// TIA Portal V21 export
// export: Created 2026-11-11T00:47:22.4274178Z, ExportSetting WithDefaults, DisplayName Totally Integrated Automation Portal, DisplayVersion V21 Update 3, DisplayName STEP 7 Professional, DisplayVersion V21 Update 3, DisplayName STEP 7 Safety, DisplayVersion V21, DisplayName Tech WebApplication, DisplayVersion V21, DisplayName WinCC Basic/Comfort/Advanced, DisplayVersion V21 Update 3, DisplayName WinCC Unified, DisplayVersion V21 Update 3
FUNCTION_BLOCK "FB_Fbd_ex066"   // FB102, FBD
{ S7_Optimized_Access := 'TRUE' }
VERSION : 0.1
// stored: AutoNumber true, IsIECCheckEnabled false, IsRetainMemResEnabled false, MemoryReserve 100, SetENOAutomatically false, UDAEnableTagReadback false
   VAR_INPUT
      v_req : Bool;
      v_r : Bool;
      v_dp_id : HW_IOSYSTEM;
   END_VAR
   VAR_OUTPUT
      v_ret_val : Int;
      v_busy : Bool;
      v_dpr : Byte;
      v_dpri : Byte;
   END_VAR
BEGIN

REGION Network 1: DP_TOPOL - Determine topology for DP master system
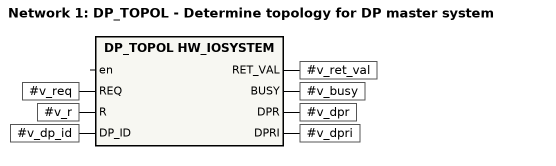
   #v_ret_val := DP_TOPOL(REQ := #v_req,
                          R := #v_r,
                          DP_ID := #v_dp_id,
                          BUSY => #v_busy,
                          DPR => #v_dpr,
                          DPRI => #v_dpri);
END_REGION
END_FUNCTION_BLOCK
